// TIA Portal V20 export
// export: Created 2026-10-19T18:06:31.7293889Z, ExportSetting WithDefaults, DisplayName Totally Integrated Automation Portal, DisplayVersion V20 Update 6, DisplayName TIA Portal Openness, DisplayVersion V20 Update 6, DisplayName TIA Portal Version Control Interface, DisplayVersion V20 Update 6, DisplayName SINAMICS Startdrive Advanced, DisplayVersion V20 SP1, DisplayName SINAMICS Startdrive G130, G150, S120, S150, SINAMICS MV, G220, S200, S210, DisplayVersion V20 SP1, DisplayName SINAMICS Startdrive G110M, G120, G120C, G120D, G120P, G115D, DisplayVersion V20 SP1, DisplayName STEP 7 Professional, DisplayVersion V20 Update 6, DisplayName STEP 7 Safety, DisplayVersion V20 Update 2, DisplayName WinCC Basic/Comfort/Advanced, DisplayVersion V20 Update 6, DisplayName WinCC Unified, DisplayVersion V20 Update 6
FUNCTION_BLOCK "SAI_IND_WriteDigitalOutputs"   // FB3, LAD
{ S7_Optimized_Access := 'FALSE' }
VERSION : 0.1
// stored: AutoNumber true, IsIECCheckEnabled false, SetENOAutomatically false, UDAEnableTagReadback false
   VAR_INPUT
      ID : HW_IO;
      Output1 : Bool;
      Output2 : Bool;
      Output3 : Bool;
      Output4 : Bool;
      Output5 : Bool;
   END_VAR
   VAR_OUTPUT
      Done : Bool;
      Error : Bool;
   END_VAR
   VAR_IN_OUT
      Write : Bool;
   END_VAR
   VAR DB_SPECIFIC
      "Step" : Int;
      Writing : Bool;
      WritePre : Bool;
      BusyNTrig : Bool;
   END_VAR
   VAR
      WRREC { S7_SetPoint := 'True'} : WRREC;
   END_VAR
   VAR_TEMP
      Length : UInt;
   END_VAR
   VAR_TEMP   // added for the SCL form of the ladder/FBD networks
      _w1 : Bool;
      _w2 : Bool;
   END_VAR
BEGIN

REGION Network 1: Initialization
   // Initializes DONE and ERROR output bits
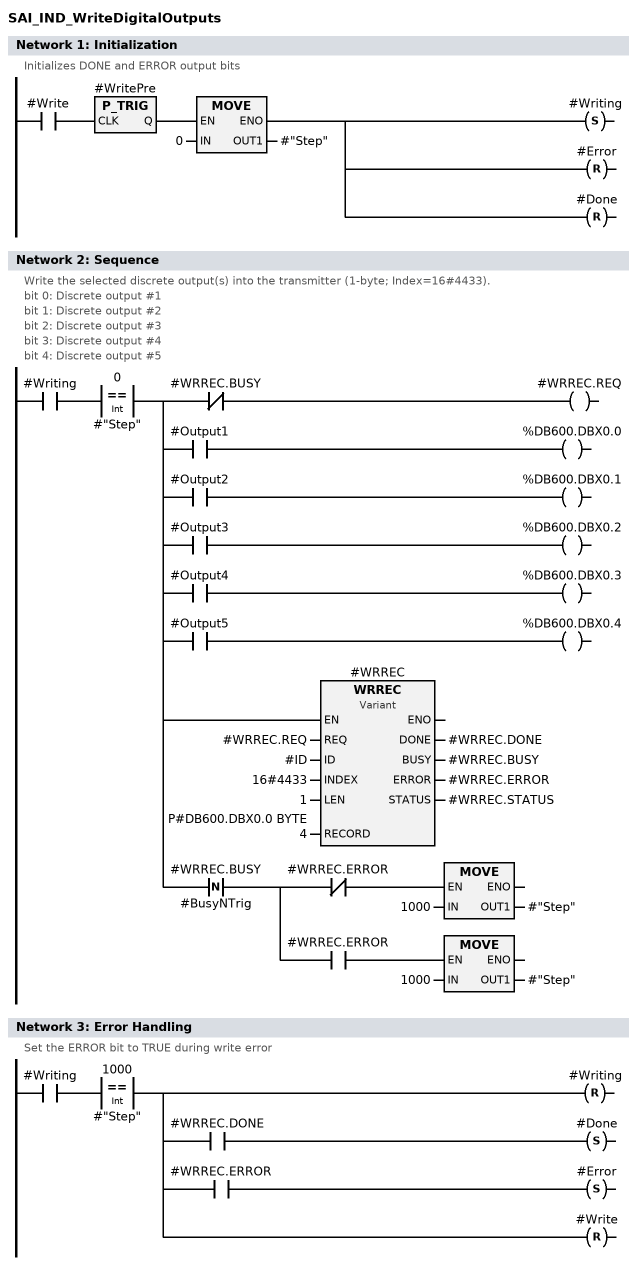
   RUNG wire#powerrail
      Contact( #Write )
      P_Trig( #WritePre )
      { S7_GenerateENO := "TRUE" } Move(in := 0, out1 => #"Step")
      wire#w1
      S_Coil( #Writing )
   END_RUNG
   RUNG wire#w1
      R_Coil( #Error )
   END_RUNG
   RUNG wire#w1
      R_Coil( #Done )
   END_RUNG
   // the same network as SCL:
   // ENO of a box is taken as its EN; it also drops when the box reports an error
   #_w1 := #Write AND NOT #WritePre;   // rising edge
   #WritePre := #Write;
   IF #_w1 THEN
       #"Step" := 0;
       #Writing := TRUE;
       #Error := FALSE;
       #Done := FALSE;
   END_IF;
END_REGION

REGION Network 2: Sequence
   // Write the selected discrete output(s) into the transmitter (1-byte; Index=16#4433).
   // bit 0: Discrete output #1
   // bit 1: Discrete output #2
   // bit 2: Discrete output #3
   // bit 3: Discrete output #4
   // bit 4: Discrete output #5
   RUNG wire#powerrail
      Contact( #Writing )
      { S7_Templates := "SrcType := Int" } EQ_Contact(in1 := 0, in2 := #"Step")
      wire#w1
      I_Contact( #WRREC.BUSY )
      Coil( #WRREC.REQ )
   END_RUNG
   RUNG wire#w1
      Contact( #Output1 )
      Coil( %DB600.DBX0.0 )
   END_RUNG
   RUNG wire#w1
      Contact( #Output2 )
      Coil( %DB600.DBX0.1 )
   END_RUNG
   RUNG wire#w1
      Contact( #Output3 )
      Coil( %DB600.DBX0.2 )
   END_RUNG
   RUNG wire#w1
      Contact( #Output4 )
      Coil( %DB600.DBX0.3 )
   END_RUNG
   RUNG wire#w1
      Contact( #Output5 )
      Coil( %DB600.DBX0.4 )
   END_RUNG
   RUNG wire#w1
      { S7_Templates := "[ptr_type := Variant, id_type := HW_IO, index_type := DInt, len_type := UInt]" } #WRREC.WRREC(REQ := #WRREC.REQ, ID := #ID, INDEX := 16#4433, LEN := 1, RECORD := P#DB600.DBX0.0 BYTE 4, DONE => #WRREC.DONE, BUSY => #WRREC.BUSY, ERROR => #WRREC.ERROR, STATUS => #WRREC.STATUS)
   END_RUNG
   RUNG wire#w1
      N_Contact(operand := #WRREC.BUSY, bit := #BusyNTrig)
      wire#w2
      I_Contact( #WRREC.ERROR )
      { S7_GenerateENO := "TRUE" } Move(in := 1000, out1 => #"Step")
   END_RUNG
   RUNG wire#w2
      Contact( #WRREC.ERROR )
      { S7_GenerateENO := "TRUE" } Move(in := 1000, out1 => #"Step")
   END_RUNG
   // the same network as SCL:
   #_w1 := #Writing AND (0 = #"Step");
   #WRREC.REQ := #_w1 AND NOT #WRREC.BUSY;
   %DB600.DBX0.0 := #_w1 AND #Output1;
   %DB600.DBX0.1 := #_w1 AND #Output2;
   %DB600.DBX0.2 := #_w1 AND #Output3;
   %DB600.DBX0.3 := #_w1 AND #Output4;
   %DB600.DBX0.4 := #_w1 AND #Output5;
   IF #_w1 THEN
       #WRREC(REQ := #WRREC.REQ,   // WRREC
              ID := #ID,
              INDEX := 16#4433,
              LEN := 1,
              RECORD := P#DB600.DBX0.0 BYTE 4,
              DONE => #WRREC.DONE,
              BUSY => #WRREC.BUSY,
              ERROR => #WRREC.ERROR,
              STATUS => #WRREC.STATUS);
   END_IF;
   #_w2 := #_w1 AND NOT #WRREC.BUSY AND #BusyNTrig;   // falling edge of #WRREC.BUSY
   #BusyNTrig := #WRREC.BUSY;
   IF #_w2 AND NOT #WRREC.ERROR THEN #"Step" := 1000; END_IF;
   IF #_w2 AND #WRREC.ERROR THEN #"Step" := 1000; END_IF;
END_REGION

REGION Network 3: Error Handling
   // Set the ERROR bit to TRUE during write error
   RUNG wire#powerrail
      Contact( #Writing )
      { S7_Templates := "SrcType := Int" } EQ_Contact(in1 := 1000, in2 := #"Step")
      wire#w1
      R_Coil( #Writing )
   END_RUNG
   RUNG wire#w1
      Contact( #WRREC.DONE )
      S_Coil( #Done )
   END_RUNG
   RUNG wire#w1
      Contact( #WRREC.ERROR )
      S_Coil( #Error )
   END_RUNG
   RUNG wire#w1
      R_Coil( #Write )
   END_RUNG
   // the same network as SCL:
   #_w1 := #Writing AND (1000 = #"Step");
   IF #_w1 THEN #Writing := FALSE; END_IF;
   IF #_w1 AND #WRREC.DONE THEN #Done := TRUE; END_IF;
   IF #_w1 AND #WRREC.ERROR THEN #Error := TRUE; END_IF;
   IF #_w1 THEN #Write := FALSE; END_IF;
END_REGION
END_FUNCTION_BLOCK
